//{attribute 'qualified_only'}
VAR_GLOBAL	
	fbPis			: ARRAY[0..E_Pis_Name.last] OF FB_Piston;
	stPis			: ARRAY[0..E_Pis_Name.last] OF ST_Piston;
	arPisName		: ARRAY[0..E_Pis_Name.last] OF ST_Piston_SelectionList;
	

	iPis_sel		: INT:=1;
	
	arPisNameList	: ARRAY[0..E_Pis_Name.last] OF STRING(12);
	ePisNameList	: E_Pis_Name;

	fbPis_U_L		: ARRAY[0..E_Pis_Name.last] OF FB_Piston_U_L;
	stPis_U_L		: ARRAY[0..E_Pis_Name.last] OF ST_Piston_U_L;

	
END_VAR

VAR_GLOBAL PERSISTENT
	stPisSetting	: ARRAY[0..E_Pis_Name.last] OF ST_Piston_Setting_Param;
END_VAR

VAR_GLOBAL CONSTANT
	C_MAX_Pistons		: INT:=E_Pis_Name.last;
	//C_MAX_Pistons_Exist	: INT:=51;	
END_VAR

(* stored: Version 1.1.0.1, ProductVersion 3.1.4024.13
   GVL g_Piston: Id {79a36863-b789-4b6c-b41a-a21efa0eb605} *)
